// TIA Portal V21 export
// export: Created 2026-11-10T07:35:17.2244837Z, ExportSetting WithDefaults, DisplayName Totally Integrated Automation Portal, DisplayVersion V21 Update 3, DisplayName STEP 7 Professional, DisplayVersion V21 Update 3, DisplayName STEP 7 Safety, DisplayVersion V21, DisplayName Tech WebApplication, DisplayVersion V21, DisplayName WinCC Basic/Comfort/Advanced, DisplayVersion V21 Update 3, DisplayName WinCC Unified, DisplayVersion V21 Update 3
FUNCTION_BLOCK "FB_Lad_ex128"   // FB101, LAD
{ S7_Optimized_Access := 'TRUE' }
VERSION : 0.1
// stored: AutoNumber true, IsIECCheckEnabled false, IsRetainMemResEnabled false, MemoryReserve 100, SetENOAutomatically false, UDAEnableTagReadback false
   VAR_INPUT
      v_laddr : HW_IOSYSTEM;
      v_station_nr : UInt;
   END_VAR
   VAR_OUTPUT
      v_done : Bool;
      v_busy : Bool;
      v_error : Bool;
      v_len : DInt;
      v_status : Word;
   END_VAR
   VAR_IN_OUT
      v_data : Array[0..99] of Byte;
   END_VAR
   VAR
      inst { S7_SetPoint := 'True'} : Get_Name;
   END_VAR
BEGIN

REGION Network 1: GET_NAME - Read out name of an IO device or a DP slave
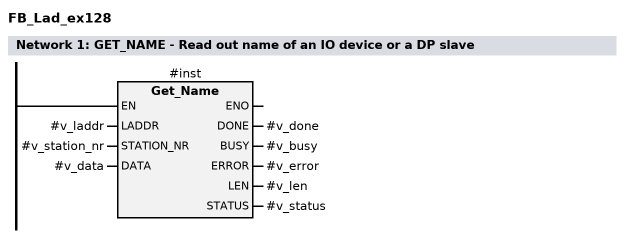
   RUNG wire#powerrail
      #inst.Get_Name(LADDR := #v_laddr, STATION_NR := #v_station_nr, DATA := #v_data, DONE => #v_done, BUSY => #v_busy, ERROR => #v_error, LEN => #v_len, STATUS => #v_status)
   END_RUNG
   // the same network as SCL:
   #inst(LADDR := #v_laddr,   // Get_Name
         STATION_NR := #v_station_nr,
         DATA := #v_data,
         DONE => #v_done,
         BUSY => #v_busy,
         ERROR => #v_error,
         LEN => #v_len,
         STATUS => #v_status);
END_REGION
END_FUNCTION_BLOCK
